Fanuc KAREL source: KT00652.KL

PROGRAM KT00652
%NOLOCKGROUP
VAR
  P1: POSITION
  P2: POSITION
  OUT: INTEGER
BEGIN
  OUT = NOT P1
END KT00652
